(*
    Legacy MPA actuator block of the kfe and lfe projects, kept as it behaved. It is not the
    library actuator: it commands itself to match a limit switch it finds active, takes its
    fast fault name from sName, and its MPS rule follows the commanded direction.
    FB_PneumaticActuator is the library block for new devices.
    The limit switch state, the insert and retract exclusion and the output timeout come from
    FB_PneumaticCore, which FB_PneumaticActuator uses as well. bEnableFF FALSE skips the fast fault.
*)
FUNCTION_BLOCK FB_MPA
VAR_INPUT
    (*EPS Interlock Bits*)
    ibInsertOK: BOOL;
    ibRetractOK: BOOL;
    ibPMPS_OK:BOOL;
    ibOverrideInterlock:BOOL; (*if true interlocks are ignored*)
    // Reset fault
    {attribute 'pytmc' := '
    pv: FF_Reset
    '}
    i_xReset: BOOL;
    bEnableFF: BOOL := TRUE;
END_VAR
VAR_OUTPUT
    {attribute 'pytmc' := '
    pv:
    '}
    q_stAct :  ST_MPA;
    {attribute 'pytmc' := '
    pv: MPS_FAULT
    '}
    xMPS_OK:BOOL;
    {attribute 'pytmc' := '
    pv: MOT_DONE
    '}
    xDone:Bool; // Motion is Done
END_VAR
VAR
    // Fast fault output the fault is raised on, and the name of the device in the fault
    fbFFHWO: REFERENCE TO FB_HardwareFFOutput;
    sName: STRING;

    // PMPS
    fbFF :  FB_FastFault :=(
        i_xAutoReset := TRUE,
        i_Desc := 'Device is moving',
        i_TypeCode := 16#1010
    );

    (*Init*)
    xFirstPass    :    BOOL;
    fbFSInit        :    R_TRIG;

    (* Shared behaviour of the pneumatic actuator blocks *)
    fbCore: FB_PneumaticCore;

    (* Timeouts*)
    tTimeOutDuration: TIME:= T#5S;

    (*IO*)
    i_xInsertedLS    AT%I*: BOOL;
    i_xRetractedLS    AT%I*: BOOL;
    q_xInsert_DO    AT%Q*: BOOL;
    q_xRetract_DO    AT%Q*: BOOL;

    (* Reset Triggers *)
    rtInsert: R_TRIG;
    rtRemove: R_TRIG;
END_VAR

IF NOT __ISVALIDREF(fbFFHWO) THEN
    RETURN;
END_IF

(*Initialize*)
fbFSInit( CLK := TRUE, Q => xFirstPass);
(*IO Mapping*)
UpdateIO();

IF xFirstPass THEN
    q_stAct.eState := E_PnuematicActuatorPositionState.INVALID;
    q_stAct.bRetract_SW := FALSE;
    q_stAct.bInsert_SW := FALSE;
END_IF


(* Manage States*)
// The output bits are those of the previous scan, so the timeout is reported one scan late
fbCore(
    bInLimitSwitch := q_stAct.i_bInLS,
    bOutLimitSwitch := q_stAct.i_bOutLS,
    bInsertOutput := q_stAct.q_bInsert,
    bRetractOutput := q_stAct.q_bRetract,
    tTimeout := tTimeOutDuration,
    eState => q_stAct.eState
);

(*Set the Done signal*)
xDone := (q_stAct.bRetract_SW AND q_stAct.eState=E_PnuematicActuatorPositionState.RETRACTED)
        OR (q_stAct.eState=E_PnuematicActuatorPositionState.INSERTED AND q_stAct.bInsert_SW);


(*MPS FAULT*)
(**)
xMPS_OK := (q_stAct.bRetract_SW AND i_xRetractedLS) XOR (i_xInsertedLS AND q_stAct.bInsert_SW);
//xMPS_OK := i_xRetractedLS XOR i_xInsertedLS;
//xMPS_OK := (q_stAct.eState=RETRACTED) OR (q_stAct.eState=INSERTED);
//xMPS_OK := (q_stAct.eState=RETRACTED) ;

(*PMPS PERMISSION*)

(* Reset the other command bit when one goes high *)
rtInsert(CLK:=q_stAct.bInsert_SW);
IF rtInsert.Q THEN
    q_stAct.bRetract_SW := FALSE;
END_IF
rtRemove(CLK:=q_stAct.bRetract_SW);
IF rtRemove.Q THEN
    q_stAct.bInsert_SW := FALSE;
END_IF

(* Can't have bRetract_SW and  bInsert_SW both be true*)
IF q_stAct.bInsert_SW AND q_stAct.bRetract_SW THEN
    q_stAct.bInsert_SW := FALSE;
    q_stAct.bRetract_SW := FALSE;
END_IF

(* Make the state consistent if we can *)
IF NOT (q_stAct.bRetract_SW OR q_stAct.bInsert_SW) THEN
    IF q_stAct.eState = E_PnuematicActuatorPositionState.RETRACTED THEN
        q_stAct.bRetract_SW := TRUE;
    ELSIF q_stAct.eState = E_PnuematicActuatorPositionState.INSERTED THEN
        q_stAct.bInsert_SW := TRUE;
    END_IF
END_IF

q_stAct.bRetractOK := ibRetractOK;
q_stAct.bInsertOK := ibInsertOK;

(*Actuate the device*)
q_stAct.q_bRetract := q_stAct.bRetractOK AND q_stAct.bRetract_SW;
q_stAct.q_bInsert := q_stAct.bInsertOK AND q_stAct.bInsert_SW;

IF q_stAct.q_bInsert THEN
    q_stAct.q_bRetract := FALSE;
    q_stAct.bRetract_SW:= FALSE;
ELSIF q_stAct.q_bRetract THEN
    q_stAct.q_bInsert := FALSE;
    q_stAct.bInsert_SW:= FALSE;
END_IF;

///Check moving postion timout
IF fbCore.bInsertTimedOut OR fbCore.bRetractTimedOut THEN
    q_stAct.bErrorPresent := TRUE;
END_IF

(*FAST FAULT*)
IF bEnableFF THEN
    fbFF(i_DevName := sName,
        i_xOK := xMPS_OK,
        i_xReset := i_xReset,
        io_fbFFHWO := fbFFHWO
   );
END_IF

(*Soft IO Mapping*)
UpdateIO();

(* Rebinds the fast fault output and the name. Call from the CallAfterInit of an enclosing FB. *)
METHOD CallAfterInitMPA
VAR_INPUT
    fbFFHWO : REFERENCE TO FB_HardwareFFOutput;
    sName : STRING;
END_VAR
THIS^.fbFFHWO REF= fbFFHWO;
THIS^.sName := sName;
END_METHOD

(* Stores the mandatory fast fault output and device name at instantiation. *)
METHOD FB_Init : BOOL
VAR_INPUT
    // TRUE: the retain variables are initialized (reset warm / reset cold)
    bInitRetains : BOOL;
    // TRUE: the instance will be copied to the copy code afterward (online change)
    bInCopyCode : BOOL;
    fbFFHWO : REFERENCE TO FB_HardwareFFOutput;
    sName : STRING;
END_VAR
THIS^.fbFFHWO REF= fbFFHWO;
THIS^.sName := sName;
END_METHOD

(* Insert request, the bit the IN_CMD PV writes. Settable so tests and simulation can drive it. *)
PROPERTY InsertCmd : BOOL
GET
InsertCmd := q_stAct.bInsert_SW;
END_GET
SET
q_stAct.bInsert_SW := InsertCmd;
END_SET
END_PROPERTY

(* Inserted limit switch input. Settable so tests and simulation can drive it. *)
PROPERTY InsertedLS : BOOL
GET
InsertedLS := i_xInsertedLS;
END_GET
SET
i_xInsertedLS := InsertedLS;
END_SET
END_PROPERTY

(* Retract request, the bit the OUT_CMD PV writes. Settable so tests and simulation can drive it. *)
PROPERTY RetractCmd : BOOL
GET
RetractCmd := q_stAct.bRetract_SW;
END_GET
SET
q_stAct.bRetract_SW := RetractCmd;
END_SET
END_PROPERTY

(* Retracted limit switch input. Settable so tests and simulation can drive it. *)
PROPERTY RetractedLS : BOOL
GET
RetractedLS := i_xRetractedLS;
END_GET
SET
i_xRetractedLS := RetractedLS;
END_SET
END_PROPERTY

(* Time an output may stay on without reaching its limit switch. Default 5 s. *)
PROPERTY TimeoutDuration : TIME
GET
TimeoutDuration := tTimeOutDuration;
END_GET
SET
tTimeOutDuration := TimeoutDuration;
END_SET
END_PROPERTY

(* Soft IO mapping: copies the limit switch inputs into the status struct and the outputs into the
   digital outputs. Runs at the start and end of every body scan. *)
METHOD UpdateIO
(*Inputs*)
q_stAct.i_bInLS :=  i_xInsertedLS;
q_stAct.i_bOutLS := i_xRetractedLS;

(*outputs*)
q_xInsert_DO:=q_stAct.q_bInsert;
q_xRetract_DO:=q_stAct.q_bRetract;
END_METHOD

END_FUNCTION_BLOCK

(* stored: Version 1.1.0.1
   POU FB_MPA: Id {cb866698-d8bc-42c2-8e0e-dd29cc758464}, SpecialFunc None
   Method CallAfterInitMPA: Id {1307ee02-c964-4b0d-b3e3-8107def010b9}
   Method FB_Init: Id {f8c83a0a-680d-4665-aefd-945fc7da00d9}
   Property InsertCmd: Id {8c76249c-195d-40c9-aa74-ef053317a39f}
   Get Get: Id {f8551b05-6b31-4d3e-8571-b4cc0e7e5406}
   Set Set: Id {93a94d89-250d-445c-8606-1254c4892110}
   Property InsertedLS: Id {812a1c9a-744b-4748-b834-3ccaf504cf3b}
   Get Get: Id {24e26031-df73-4459-b753-5e6ed5d716b1}
   Set Set: Id {d523f58d-fb23-45c0-83a5-b4052bfd5071}
   Property RetractCmd: Id {f2a24ff2-07ca-4d75-bfa5-6fb9c3101785}
   Get Get: Id {a2752d9d-c878-44d7-94ae-29c0a93bccfe}
   Set Set: Id {a3f15b69-d5e5-45ee-9d49-55df8cd19b28}
   Property RetractedLS: Id {c3d6a7fa-fbbb-4819-a638-2277c015090a}
   Get Get: Id {39037495-7da3-45a5-9c4a-d4862cd30ceb}
   Set Set: Id {7352f6e5-19bf-4f83-948d-b8828a446ef5}
   Property TimeoutDuration: Id {b37cc1cf-4759-4e5b-a187-d914a7d82ad9}
   Get Get: Id {8d63bb8f-9a31-436d-838b-caf58db4d421}
   Set Set: Id {c58afb99-00c5-43c2-8286-8f44840ada8f}
   Method UpdateIO: Id {57068de5-6c7f-4be2-94ad-5467e24dfe72} *)
